(* IEC 61131-3 sources: CodesysTools/tests/expected, 17 files *)

(* ---- naming_noprefix.st ---- *)
//{attribute 'noprefix'}
{attribute 'pack_mode' := '1'}
TYPE tMbUnion :
UNION
    b   : tMbState;  //For Bit Access
    dw  : DWord;     //For DoubleWord Access
    w2  : Word;
    Raw : Int;
    foo : Int;
END_UNION
END_TYPE

(* ---- naming_union.st ---- *)
{attribute 'pack_mode' := '1'}
TYPE tMbUnion :
UNION
    b   : tMbState;  //For Bit Access
    dw  : DWord;     //For DoubleWord Access
    w2  : Word;
    Raw : Int;
    foo : Int;
END_UNION
END_TYPE

(* ---- decl_init.st ---- *)
FUNCTION_BLOCK FB_X
VAR
    sValve             : tValve
        (
         bOpen         := True,
         iMax          := 10,
         rGain         := 1.5
         );  // valve
    sb                 : Bool;
    sName              : String(80) := 'x';
{attribute 'a'} sOther : tOther :=
        (
         iA            := 1,
         iB            := 2
         );
    saArr              : Array[1..2] Of Int := [1, 2];
END_VAR
sb                     := True;

(* ---- general.st ---- *)
FUNCTION_BLOCK fb_Motor EXTENDS fb_Base
VAR_INPUT
    bStart             : Bool;                        // start command
    bStop              : Bool := False;               // stop
    nSpeedSetpoint     : Int;
END_VAR
VAR
    tonDelay           : TON;
    aBuffer            : Array[1..10] Of Real;
    sName              : String(80) := 'Motor $'A$'';
    iState             : Int;
    dtStart            : DT := DT#2024-01-01-12:30:00;
    pIn AT %IX0.1      : Bool;
END_VAR

(* main logic *)
If bStart And Not bStop Then
    iState             := 1;
ElsIf bStop Then
    iState             := 0;
Else
    x                  := -5 + y * (3 - z);
End_If

Case iState Of
    0:
        tonDelay
            (
             IN        := False,
             PT        := T#2S
             );
    1, 2: tonDelay(IN := True,
            PT         := T#5s);
        If tonDelay.Q Then
            iState     := E_State#Running;
        End_If
    -1:;
Else
    iState             := 0;
End_Case

For i := 1 To 10 By 1 Do
    aBuffer[i]         := Int_To_Real(i) * 1.5E3;
End_For
Repeat
    i                  := i + 1;
Until i > 5
End_Repeat;
END_FUNCTION_BLOCK

TYPE ST_Data :
STRUCT
    a                  : Int;                         // first
    longName           : LReal := 1.0;
END_STRUCT
END_TYPE

PROGRAM Main
VAR
    i                  : Int;                         // loop counter
    rTemperatureActual : Real := 20.5;                // measured
    bAlarm             : Bool;
END_VAR
i                      := 0;                          // reset
rTemperatureActual     := rTemperatureActual + 0.1;
bAlarm                 := rTemperatureActual > 80.0;  // high temp
THIS^.x                := 1;
END_PROGRAM

(* ---- general.upper.st ---- *)
FUNCTION_BLOCK fb_Motor EXTENDS fb_Base
VAR_INPUT
    bStart             : BOOL;                        // start command
    bStop              : BOOL := FALSE;               // stop
    nSpeedSetpoint     : INT;
END_VAR
VAR
    tonDelay           : TON;
    aBuffer            : ARRAY[1..10] OF REAL;
    sName              : STRING(80) := 'Motor $'A$'';
    iState             : INT;
    dtStart            : DT := DT#2024-01-01-12:30:00;
    pIn AT %IX0.1      : BOOL;
END_VAR

(* main logic *)
IF bStart AND NOT bStop THEN
    iState             := 1;
ELSIF bStop THEN
    iState             := 0;
ELSE
    x                  := -5 + y * (3 - z);
END_IF

CASE iState OF
    0:
        tonDelay
            (
             IN        := FALSE,
             PT        := T#2S
             );
    1, 2: tonDelay(IN := TRUE,
            PT         := T#5s);
        IF tonDelay.Q THEN
            iState     := E_State#Running;
        END_IF
    -1:;
ELSE
    iState             := 0;
END_CASE

FOR i := 1 TO 10 BY 1 DO
    aBuffer[i]         := Int_To_Real(i) * 1.5E3;
END_FOR
REPEAT
    i                  := i + 1;
UNTIL i > 5
END_REPEAT;
END_FUNCTION_BLOCK

TYPE ST_Data :
STRUCT
    a                  : INT;                         // first
    longName           : LREAL := 1.0;
END_STRUCT
END_TYPE

PROGRAM Main
VAR
    i                  : INT;                         // loop counter
    rTemperatureActual : REAL := 20.5;                // measured
    bAlarm             : BOOL;
END_VAR
i                      := 0;                          // reset
rTemperatureActual     := rTemperatureActual + 0.1;
bAlarm                 := rTemperatureActual > 80.0;  // high temp
THIS^.x                := 1;
END_PROGRAM

(* ---- naming.st ---- *)
VAR_GLOBAL
    gbAlarm          : Bool;
    bAlarm2          : Bool;
    iStart AT %IX0.0 : Bool;
    ibStop AT %IX0.1 : Bool;
    qbLamp AT %QX0.0 : Bool;
END_VAR
VAR_GLOBAL CONSTANT
    gciMax           : Int := 10;
    MAX_N            : Int := 5;
END_VAR
FUNCTION_BLOCK fbMotor
VAR_INPUT
    ibReset          : Bool;
    nSpeed           : Int;
    ixEnable, bRun   : Bool;
    iAxis            : ST_Axis;
END_VAR
VAR_OUTPUT
    qrSpeed          : Real;
    qlrPos           : LReal;
END_VAR
VAR_IN_OUT
    iqData           : ST_Data;
END_VAR
VAR
    sbReset          : Bool;
    tonDelay         : TON;
    sTimer           : TON;
    aBuf             : Array[1..10] Of Real;
    srBuf2           : Array[1..10] Of Real;
    sudiCount        : UDInt := 0;
    sString          : String(80);
    ssName           : String(80);
    sdtStamp         : DT;
END_VAR
VAR CONSTANT
    ciLimit          : Int := 3;
END_VAR
VAR_TEMP
    ttElapsed        : Time;
    tData            : ST_Data;
END_VAR
END_FUNCTION_BLOCK
FUNCTION fcAdd : Int
VAR
    tiX              : Int;
    siY              : Int;
END_VAR
END_FUNCTION
TYPE ST_Data :
STRUCT
    bOk              : Bool;
    rVal             : Real;
    value            : Int;
    Sub              : ST_Sub;
END_STRUCT
END_TYPE

(* ---- naming_block_skip.st ---- *)
TYPE tA :
STRUCT  //{attribute 'noprefix'}
    Alpha   : Int;
    Beta    : Bool;
END_STRUCT
END_TYPE
TYPE tB :
STRUCT
    Gamma   : Int;
END_STRUCT
END_TYPE
FUNCTION_BLOCK FB_X
VAR     (* {attribute 'noprefix'} *)
    Free    : Int;
END_VAR
VAR
    Checked : Int;
END_VAR
END_FUNCTION_BLOCK

(* ---- naming_prefixes.st ---- *)
FUNCTION_BLOCK FB_T
VAR
    kMaxSize : Int := 3;
    vSpeed   : Real;
    mValue   : Bool;
    mode     : Int;
    kmax     : Int;
    m        : Int;
    sbOk     : Bool;
    sb2Valve : Bool;
    sbValve2 : Bool;
    k2Max    : Int;
    sb_x     : Bool;
    k        : Int;
    k_1      : Int;
    v        : Int;
    smRot    : Real;
    tmRot    : Real;
    svPos    : Real;
    tvPos2   : Real;
    tmp      : Real;
    gmRot    : Real;
END_VAR
END_FUNCTION_BLOCK

(* ---- naming_types.st ---- *)
FUNCTION_BLOCK FB_T
VAR
    Start : TOD;
    Data  : ST_Data;
    aData : Array[0..3] Of ST_Data;
    Other : ST_Other;
    Flag  : Bool;
END_VAR
END_FUNCTION_BLOCK

(* ---- region_attributes.st ---- *)
FUNCTION_BLOCK fb_Motor
VAR_INPUT
    bStart                               : Bool;           // start command
{attribute 'hide'} bInternalFlagLongName : Bool := False;  // stop
{attribute 'hide'} nCnt                  : LInt;
END_VAR
VAR_OUTPUT
    x                                    : LReal;          // out
END_VAR
REGION Motor If control
    If bStart Then
        iState                           := 1;             // run
    ElsIf bStop Then
        iCounterValue                    := 0;
    Else
        x                                := -5;
    End_If
END_REGION
For i := 1 To 10 Do
    aBuffer[i]                           := i;             // fill
End_For
END_FUNCTION_BLOCK

(* ---- spelling.st ---- *)
// This valve is wrong, the wrod is spelled wrong
(* Valves and unhappy workers check the lines *)
FUNCTION_BLOCK FB_Valve
VAR
    sbOpen    : Bool;   // The valve colour: a PLC flag with a mispelling
    sbValveOk : Bool;   // valvs of London and tMbState and sValve
END_VAR
// sbOpen := TRUE;  commented out code is skipped
// See https://example.com/wrodd and file.txt for details
sbOpen        := True;  // Worke it, e.g. unworkers and valveed
(* Multi
   line commment
   second: chek the line *)
// {attribute 'noprefix'}
// arbeidsbord og ventilbord, løs og ære, feilstavet ventilbrod
END_FUNCTION_BLOCK

(* ---- terminal_codes.st ---- *)
FUNCTION_BLOCK FB_Valve
VAR_INPUT
    R         : Bool;
    BA1       : Bool;
    XE        : Bool;
    START_CMD : Bool;
    BZ        : Bool;
    QA        : Bool;
    Start     : Bool;
    ibReset   : Bool;
END_VAR
VAR_OUTPUT
    YH        : Bool;
    qbOpen    : Bool;
END_VAR
VAR
    START     : Bool;
END_VAR
END_FUNCTION_BLOCK

(* ---- calls.align40.st ---- *)
PROGRAM Main
VAR
    sTimer                             : TON;
    sbStart                            : Bool;
    sbDone                             : Bool;
    stElapsed                          : Time;
    srX                                : Real;
END_VAR
sbStart                                := True;
sTimer
    (
     IN                                := sbStart,
     PT                                := T#5S,  // time
     Q                                 => sbDone,
     ET                                => stElapsed
     );                                          // done
If sbStart Then
    aFb[1].Run
        (
         Execute                       := True
         );
    srX                                := Limit(0.0, srX, 10.0);
    F_Calc(srX);
End_If
srX                                    := a +
F(b := 1);
sTimer
    (
     // comment line
     IN                                := sbStart
     );
END_PROGRAM

(* ---- calls.preserve.st ---- *)
PROGRAM Main
VAR
    sTimer    : TON;
    sbStart   : Bool;
    sbDone    : Bool;
    stElapsed : Time;
    srX       : Real;
END_VAR
sbStart       := True;
sTimer(IN := sbStart, PT := T#5S,           // time
    Q         => sbDone, ET => stElapsed);  // done
If sbStart Then
    aFb[1].Run(Execute := True);
    srX       := Limit(0.0, srX, 10.0);
    F_Calc(srX);
End_If
srX           := a +
F(b := 1);
sTimer(
    // comment line
    IN        := sbStart);
END_PROGRAM

(* ---- calls.st ---- *)
PROGRAM Main
VAR
    sTimer       : TON;
    sbStart      : Bool;
    sbDone       : Bool;
    stElapsed    : Time;
    srX          : Real;
END_VAR
sbStart          := True;
sTimer
    (
     IN          := sbStart,
     PT          := T#5S,  // time
     Q           => sbDone,
     ET          => stElapsed
     );                    // done
If sbStart Then
    aFb[1].Run
        (
         Execute := True
         );
    srX          := Limit(0.0, srX, 10.0);
    F_Calc(srX);
End_If
srX              := a +
F(b := 1);
sTimer
    (
     // comment line
     IN          := sbStart
     );
END_PROGRAM

(* ---- functions.st ---- *)
PROGRAM P
VAR
    sR : LReal;
END_VAR
sR     := Abs(x) + Sin(y) + Int_To_Real(i) + To_Int(r) + Max(a, b) + st.Len + Limit(0, a, 5);
sR     := stX.max;
sR     := LTime_To_LReal(a) + To_DWord(c) + Trunc_Int(d) + TOD_To_Time(f);

(* ---- typed_literals.st ---- *)
PROGRAM P
VAR
    sT : LTime := LTime#1s;
    sB : Int := Int#5;
END_VAR
sT     := TOD#12:00:00; sB := 16#FF; sT := T#5s; sT := DInt#3;
